Staubli VAL3: physicalIO.pgx

program physicalIO()
// Isma structure adapted to Level 2; taught joints, bounded cycles and shared IO modes.
begin
  // ============================================================
  // SENSORES Y ALIMENTADOR DEL LEVEL 2
  // ============================================================
  // Solo se crea en fisico. En simulacion los sensores se editan a mano.
  // La pinza usa open/close con valve1; NO escribir valve1 aqui.
  while true
    cylinderPresent = io:bIn2 == true
    feederExtended = io:bIn14 == true
    feederRetracted = io:bIn15 == true
    io:bOut10 = feederExtend
    ioReady = true
    delay(0.01)
  endWhile
end
